(* IEC 61131-3 sources: avi-aoi-management/scripts/ai-eval/ngau-nhien/kho/st-tt8-doc-tang-giam/khung/src, 1 file *)

(* ---- DocTangGiam.st ---- *)
FUNCTION_BLOCK DocTangGiam
VAR_INPUT
    DICH : REAL;
    TOC_DO_TANG : REAL;
    TOC_DO_GIAM : REAL;
    BAT : BOOL;
END_VAR
VAR_OUTPUT
    RA : REAL;
    DA_TOI : BOOL;
END_VAR
    (* TODO: cài đặt theo đề bài *)
    RA := 0.0;
END_FUNCTION_BLOCK
